// One stop per axis and stop transaction (#108), and the transaction is only settled when it is really over (#98).
// FB_TelescopeControl._StopTelescope calls the body while it stops the axes (request logic); Monitor() runs every
// scan and decides when the stop has settled: every axis that was sent a stop has reported Done, the telescope is at
// rest, and no axis has been locked for motion commands (MC_Stop, StateDWord bit 29) for 3 scans. A transaction is
// started with Begin(). A transaction that has not settled 30 s after Begin() (an axis never reports Done: its stop was
// never allowed, or the Done was lost) is released once the telescope is at rest, without the Done condition (#120);
// the stop is not sent again (the retrigger of #108 is gone). The capture of 2026-10-19 showed StandStill TRUE for one scan before the stop takes hold
// (bStopped alone released the home too early, HA error 17135). Pure logic (no axis access), tested offline in
// IAG50cmTests (#120, #98).
FUNCTION_BLOCK FB_StopTransaction
VAR_INPUT
	nTimeDivisor	: UDINT := 1;	// test seam: divides the 30 s timeout (FB_TelescopeControl.nTimeDivisor); production leaves it at 1
	bHaStandStill	: BOOL;		// HA axis at standstill (a running MC_Stop reports FALSE)
	bDecStandStill	: BOOL;
END_VAR
VAR_OUTPUT
	bStopHa			: BOOL;		// TRUE in the one scan in which the HA axis is to be sent its stop
	bStopDec		: BOOL;
	bFinished		: BOOL;		// the stop has settled: release both stop requests, the stop is done
	bActive			: BOOL;		// a transaction was begun and has not settled yet (homes and restarts wait for it)
	bTimedOut		: BOOL;		// #120: TRUE in the one scan in which the transaction passed 30 s without settling
	bHaNoDone		: BOOL;		// #120: at that moment HA was sent a stop and had not reported Done (latched until Begin/Cancel)
	bDecNoDone		: BOOL;
	bReleasedByTimeout	: BOOL;	// #120: TRUE in the one scan in which the transaction settled without a Done of a requested axis
END_VAR
VAR
	bHaStopRequested	: BOOL;		// the HA axis was sent its stop in this transaction, never again
	bDecStopRequested	: BOOL;
	bHaDone				: BOOL;		// the HA axis reported StopDone in this transaction
	bDecDone			: BOOL;
	nClearScans			: UINT;		// consecutive scans without a motion lock
	bAtRest				: BOOL;		// bStopped as seen by the last Monitor() call
	tonTimeout			: FB_TimeoutTimer;	// #120: 30 s from Begin()
	bExpired			: BOOL;		// #120: the transaction passed 30 s; the Done condition is waived from now on
END_VAR
VAR CONSTANT
	nSettleScans		: UINT := 3;	// 30 ms at the 10 ms task
	tTimeout			: TIME := T#30S;	// #120: the stop command timeout of FB_TelescopeControl (#40: a stop from slew speed takes about 4 s)
END_VAR

bStopHa := FALSE;
bStopDec := FALSE;

IF NOT bHaStopRequested AND NOT bHaStandStill THEN
	bStopHa := TRUE;
	bHaStopRequested := TRUE;
END_IF

IF NOT bDecStopRequested AND NOT bDecStandStill THEN
	bStopDec := TRUE;
	bDecStopRequested := TRUE;
END_IF

// settled (or no transaction running, as before #98): finished as soon as the telescope is at rest
bFinished := NOT bActive AND bAtRest;

// Start a new stop transaction: each axis may be sent one stop again.
METHOD Begin
bHaStopRequested := FALSE;
bDecStopRequested := FALSE;
bHaDone := FALSE;
bDecDone := FALSE;
nClearScans := 0;
bExpired := FALSE;
bHaNoDone := FALSE;
bDecNoDone := FALSE;
tonTimeout(IN := FALSE, PT := tTimeout, nDivisor := nTimeDivisor);
bActive := TRUE;
END_METHOD

// Call every scan. A transaction settles when every axis that was sent a stop has reported Done (a disabled axis
// counts as done), the telescope is at rest and no enabled axis has been locked for nSettleScans scans.
// A running calibration sweep (bHaHoming / bDecHoming) is aborted first (#113).
// #120: 30 s after Begin() a transaction that has not settled stops waiting for the Done of the axes (bTimedOut); it
// settles as soon as the telescope is at rest, no axis has been locked for nSettleScans scans and no sweep homing runs
// (bReleasedByTimeout if an axis never reported Done).
METHOD Monitor
VAR_INPUT
	bStopped		: BOOL;		// the whole telescope is at rest
	bHaEnabled		: BOOL;
	bDecEnabled		: BOOL;
	bHaStopDone		: BOOL;		// StopDone pulse of the HA axis
	bDecStopDone	: BOOL;
	bHaLocked		: BOOL;		// MotionCommandsLocked (StateDWord bit 29) of the HA axis
	bDecLocked		: BOOL;
	bHaHoming		: BOOL;		// #113: the calibration sweep of the axis is still running or being aborted (FB_LatchHome.Busy)
	bDecHoming		: BOOL;
END_VAR
bTimedOut := FALSE;
bReleasedByTimeout := FALSE;

IF bHaStopDone THEN
	bHaDone := TRUE;
END_IF
IF bDecStopDone THEN
	bDecDone := TRUE;
END_IF

IF (bHaEnabled AND bHaLocked) OR (bDecEnabled AND bDecLocked) THEN
	nClearScans := 0;
ELSIF nClearScans < nSettleScans THEN
	nClearScans := nClearScans + 1;
END_IF

bAtRest := bStopped;

tonTimeout(IN := bActive, PT := tTimeout, nDivisor := nTimeDivisor);
IF bActive AND tonTimeout.Q AND NOT bExpired THEN
	bExpired := TRUE;
	bTimedOut := TRUE;
	bHaNoDone := bHaStopRequested AND NOT bHaDone AND bHaEnabled;
	bDecNoDone := bDecStopRequested AND NOT bDecDone AND bDecEnabled;
END_IF

IF bActive
	AND bStopped
	AND (NOT bHaStopRequested OR bHaDone OR NOT bHaEnabled OR bExpired)
	AND (NOT bDecStopRequested OR bDecDone OR NOT bDecEnabled OR bExpired)
	AND nClearScans >= nSettleScans
	AND NOT bHaHoming AND NOT bDecHoming THEN
	bActive := FALSE;
	bReleasedByTimeout := bExpired AND
		((bHaStopRequested AND NOT bHaDone AND bHaEnabled) OR (bDecStopRequested AND NOT bDecDone AND bDecEnabled));
END_IF
END_METHOD

// Forget a running transaction (error, reset): nothing waits for it any more.
METHOD Cancel
bActive := FALSE;
bExpired := FALSE;
bHaNoDone := FALSE;
bDecNoDone := FALSE;
tonTimeout(IN := FALSE, PT := tTimeout, nDivisor := nTimeDivisor);
END_METHOD

END_FUNCTION_BLOCK

(* stored: Version 1.1.0.1, ProductVersion 3.1.4024.15
   POU FB_StopTransaction: Id {5a92265e-6a39-40df-a29a-dd046a1da95a}, SpecialFunc None
   Method Begin: Id {531e9405-351a-49d1-a616-de19bbf299ad}
   Method Monitor: Id {48fd0ac6-2d4c-4c9d-a1b6-2c75f44edc09}
   Method Cancel: Id {738c7907-e27e-47d5-be26-0ad891eee46f} *)
